Universal Robots URScript: T003_qwen2.5-coder_32b-instruct-q4_0_baseline_rep1.urscript

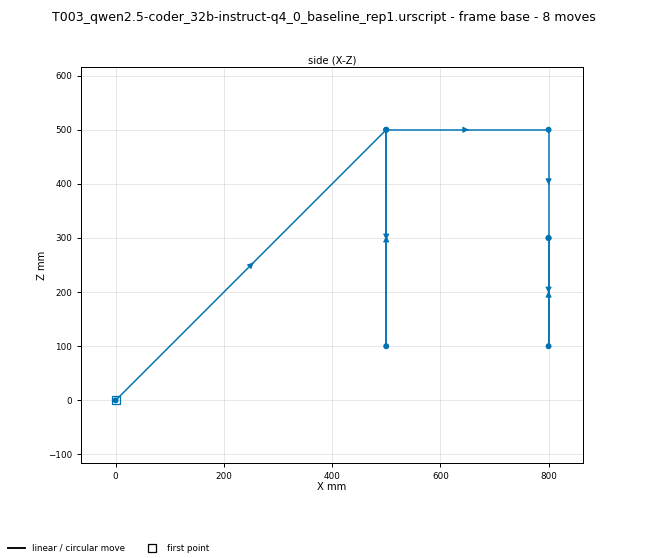
[picture p0: tool path of T003_qwen2.5-coder_32b-instruct-q4_0_baseline_rep1.urscript in frame base, 8 of 8 moves have a stored position in this frame; points joined in program order, loops and branches not executed]
# Home position
movej(p[0.0, -1.5708, 0.0, -1.5708, 0.0, 0.0], a=1.2, v=1.2, t=0, r=0)

# Approach conveyor pick — above
movel(p[0.5, -1.5708, 0.5, -1.5708, 0.0, 0.0], a=1.2, v=0.25, t=0, r=0)

# Descend to pick
movel(p[0.5, -1.5708, 0.1, -1.5708, 0.0, 0.0], a=1.2, v=0.1, t=0, r=0)

# Lift from conveyor
movel(p[0.5, -1.5708, 0.5, -1.5708, 0.0, 0.0], a=1.2, v=0.2, t=0, r=0)

# Transit to pallet position (0,0)
movel(p[0.8, -1.5708, 0.5, -1.5708, 0.0, 0.0], a=1.2, v=0.28, t=0, r=0)

# Approach pallet position (0,0) — above
movel(p[0.8, -1.5708, 0.3, -1.5708, 0.0, 0.0], a=1.2, v=0.25, t=0, r=0)

# Descend to place
movel(p[0.8, -1.5708, 0.1, -1.5708, 0.0, 0.0], a=1.2, v=0.1, t=0, r=0)

# Lift from pallet
movel(p[0.8, -1.5708, 0.3, -1.5708, 0.0, 0.0], a=1.2, v=0.2, t=0, r=0)
